Fanuc KAREL source: KA00022.KL

PROGRAM KA00022
%NOLOCKGROUP
VAR
  SRC: REAL
  DST: CONFIG
BEGIN
  SRC = 2.0
  DST = SRC
END KA00022
